Fanuc KAREL source: kt00017.KL

-- PROVISIONAL review KL for V1013-1; original PC SHA256 8b0d2d2d704a60a10853bd3ef0c973eb560983ff60e78fe43a907ed21f4926f4
-- Incomplete behavior may be omitted. Consult companion uncertainty JSON. Do not deploy.
PROGRAM KT00017
%NOLOCKGROUP
VAR
  I2 : INTEGER
  OUT : INTEGER
-- UNRESOLVED_DECL Y1 type=002018
BEGIN
  -- UNRESOLVED_PC offsets 5-19; opcodes 2E,22,9D,33,B2
  -- UNRESOLVED_PC offsets 24-35; opcodes 2E,23
  -- UNRESOLVED_PC offsets 40-62; opcodes 22,9D,33,B1,21,52,23
  -- UNRESOLVED_PC offsets 67-71; opcodes 7F
END KT00017
